TYPE U_UINT16 :
UNION
	Bits : ARRAY [1..1] OF  ST_Bits;
	Num : UINT;
END_UNION
END_TYPE

(* stored: Version 1.1.0.1
   DUT U_UINT16: Id {4b67ac90-9d43-4d5c-87a7-9e985730d07c} *)
